(*
SPDX-FileCopyrightText: © 2026 Oleksandr Tiutyk <trofimich@gmail.com>
SPDX-License-Identifier: MIT
License: https://opensource.org/license/mit
*)

(*
Observes Workflow.InitializeVariables and Workflow.OnReinitVariables during FB_reinit checks.

Binds borrowed counter storage in InitializeVariables and optionally rebinds relocated counter storage in
OnReinitVariables without throwing or clearing previously assigned values.
*)

{attribute 'no_explicit_call' := 'do not call this function block directly'}
{attribute 'no_assign'}
FUNCTION_BLOCK WorkflowOnlineChangeWorkflow EXTENDS TOF_Workflow.Workflow
VAR_STAT
	// Distinct static field to avoid redeclaring inherited Workflow metadata.
	{attribute 'hide'}
	_ProbeClassName : STRING := __POUNAME();
END_VAR
VAR
	_InitialCounter : POINTER TO DINT;
	_RelocatedCounter : POINTER TO DINT;
	_UseRelocatedTarget : BOOL;
	_InitializeCount : DINT;
	_ReinitVariablesCount : DINT;
END_VAR

(* Configures the borrowed initial and relocated DINT variable storage addresses. *)
METHOD ConfigureCounterTargets
VAR_INPUT
	initialTarget : POINTER TO DINT;
	relocatedTarget : POINTER TO DINT;
END_VAR
_InitialCounter := initialTarget;
_RelocatedCounter := relocatedTarget;
_UseRelocatedTarget := FALSE;
_InitializeCount := 0;
_ReinitVariablesCount := 0;
END_METHOD

(* Enables rebinding Counter to relocatedTarget on subsequent OnReinitVariables calls. *)
METHOD EnableRelocatedRebind
_UseRelocatedTarget := TRUE;
END_METHOD

(* Binds Counter to the initial storage address when configured. *)
METHOD PROTECTED InitializeVariables
_InitializeCount := _InitializeCount + 1;

IF _InitialCounter <> 0 THEN
	BindPlcVariable(name := 'Counter', plcVariable := _InitialCounter^);
END_IF
END_METHOD

(* Counts OnReinitVariables invocations and rebinds Counter when relocated rebinding is active. *)
METHOD PROTECTED OnReinitVariables
_ReinitVariablesCount := _ReinitVariablesCount + 1;

IF _UseRelocatedTarget AND_THEN _RelocatedCounter <> 0 THEN
	TryRebindPlcVariable(name := 'Counter', plcVariable := _RelocatedCounter^);
END_IF
END_METHOD

(* Reports the number of InitializeVariables invocations observed on this workflow. *)
{attribute 'monitoring' := 'call'}
PROPERTY InitializeCount : DINT
GET
InitializeCount := _InitializeCount;
END_GET
END_PROPERTY

(* Reports the number of OnReinitVariables invocations observed on this workflow. *)
{attribute 'monitoring' := 'call'}
PROPERTY ReinitVariablesCount : DINT
GET
ReinitVariablesCount := _ReinitVariablesCount;
END_GET
END_PROPERTY

// Borrows the concrete class name. Callers must not modify it.
{attribute 'monitoring' := 'call'}
PROPERTY ClassName : REFERENCE TO STRING
GET
ClassName REF= _ProbeClassName;
END_GET
END_PROPERTY

// Borrows the compiler-initialized namespace name. Callers must not modify it.
{attribute 'monitoring' := 'call'}
PROPERTY NamespaceName : REFERENCE TO STRING
GET
// SA0006: Read-only namespace string borrowed across test tasks.
{analysis -6}
NamespaceName REF= CurrentNamespace.Name;
{analysis +6}
END_GET
END_PROPERTY

// Reports the concrete instance size in bytes.
{attribute 'monitoring' := 'call'}
PROPERTY SelfSize : ULINT
GET
SelfSize := XSIZEOF(THIS^);
END_GET
END_PROPERTY

END_FUNCTION_BLOCK

(* stored: Version 1.1.0.1
   POU WorkflowOnlineChangeWorkflow: Id {36b07a73-6955-44bd-87d6-9fb7b587aab2}, SpecialFunc None
   Method ConfigureCounterTargets: Id {39e2d875-6026-45c6-b932-2b928cf410b9}
   Method EnableRelocatedRebind: Id {c8658395-756d-4867-bf41-58f02419065e}
   Method InitializeVariables: Id {8a48dadb-775a-4bd5-a2db-8e3d8f59db04}
   Method OnReinitVariables: Id {3145991e-2e1f-47c7-9232-576c241f05ac}
   Property InitializeCount: Id {5c5c6d92-d86e-4451-9ddd-a2e995bdd19b}
   Get Get: Id {9c217bb8-eab3-488b-aab3-91c2c32eb3a5}
   Property ReinitVariablesCount: Id {379275ec-5f17-4b81-b77e-a9730af43cb3}
   Get Get: Id {5a48df0a-9a71-4a94-93db-4653c5d0cb4d}
   Property ClassName: Id {e6b1f38a-e0a8-4ff7-9472-eee5b2f5e3aa}
   Get Get: Id {52a05038-c0b0-42f8-b935-44565fa165b7}
   Property NamespaceName: Id {0210bf12-7c9a-4c25-b3cb-ce44914e8e18}
   Get Get: Id {57a853f2-e42f-491d-97be-d09aab991eaf}
   Property SelfSize: Id {cb3e169a-d8ad-4bb6-aeca-e5f44dcaa4fb}
   Get Get: Id {837dc655-d15e-4837-99c6-d669ef7be49e} *)
